(* IEC 61131-3 sources: codesys-framework/txt/application/WeVe Core (library)/60 Event/Service/FB_EventService, 4 files *)

(* ---- FB_Init.method.st ---- *)
//FB_Init is always available implicitly and it is used primarily for initialization.
//The return value is not evaluated. For a specific influence, you can also declare the
//methods explicitly and provide additional code there with the standard initialization
//code. You can evaluate the return value.
METHOD FB_Init: BOOL
VAR_INPUT
    bInitRetains: BOOL; // TRUE: the retain variables are initialized (reset warm / reset cold)
    bInCopyCode: BOOL;  // TRUE: the instance will be copied to the copy code afterward (online change)

	fbLogger 		: I_Logger;		// mag 0 zijn
END_VAR
// --- BEGIN IMPLEMENTATION ---

// Enkel referenties bewaren, geen methodes aanroepen
_fbLogger := fbLogger;

(* ---- Initialize.method.st ---- *)
// Eenmalig bij de opstart, na het registreren: alle groepen initialiseren
// (logger doorgeven, config invullen). Groepen die later registreren worden meteen geïnitialiseerd.
// TRUE = klaar.
METHOD Initialize : BOOL
VAR_INPUT
END_VAR
VAR
	i 		: INT;
END_VAR
// --- BEGIN IMPLEMENTATION ---

FOR i := 0 TO _iGroupCount - 1 DO
	IF _afbGroups[i] <> 0 THEN
		_afbGroups[i].Initialize();
	END_IF
END_FOR

_xInitialized := TRUE;
Initialize := TRUE;

(* ---- Register.method.st ---- *)
// Een EventGroup registreren. Bij de opstart, vanuit FB_Application.
// Registreren na Initialize mag ook: de groep wordt dan meteen geïnitialiseerd.
// FALSE = groep is 0, al geregistreerd, of de lijst is vol (wordt gelogd).
METHOD Register : BOOL
VAR_INPUT
	fbEventGroup 	: I_EventGroup;
END_VAR
VAR
	i 				: INT;
END_VAR

// --- BEGIN IMPLEMENTATION ---

IF fbEventGroup = 0 THEN
	Register := FALSE;
	RETURN;
END_IF

// Dubbele registratie
FOR i := 0 TO _iGroupCount - 1 DO
	IF _afbGroups[i] = fbEventGroup THEN
		Register := FALSE;
		RETURN;
	END_IF
END_FOR

// Lijst vol: nooit stil negeren
IF _iGroupCount >= cMaxGroups THEN
	IF _fbLogger <> 0 THEN
		_fbLogger.LogMessage(
			eLevel 		:= E_EventLevels.EventIsAlarm_OnlyLogLevel,
			sMessage 	:= 'FB_EventService: too many event groups, increase cMaxGroups');
	END_IF
	Register := FALSE;
	RETURN;
END_IF

_afbGroups[_iGroupCount] := fbEventGroup;
_iGroupCount := _iGroupCount + 1;

IF _xInitialized THEN
	fbEventGroup.Initialize();
END_IF

Register := TRUE;

(* ---- Reset.method.st ---- *)
// Globale reset: alle groepen resetten. Elk event beslist zelf of het mag (conditie weg).
// TRUE = geen enkel event nog actief.
METHOD Reset : BOOL
VAR_INPUT
END_VAR
VAR
	i 			: INT;
	xAllReset 	: BOOL := TRUE;
END_VAR

// --- BEGIN IMPLEMENTATION ---

FOR i := 0 TO _iGroupCount - 1 DO
	IF _afbGroups[i] <> 0 THEN
		// Reset altijd aanroepen, ook als een vorige groep al FALSE gaf
		IF NOT _afbGroups[i].Reset() THEN
			xAllReset := FALSE;
		END_IF
	END_IF
END_FOR

Reset := xAllReset;
